Fanuc KAREL source: kb00020.KL

-- PROVISIONAL review KL for V1013-1; original PC SHA256 263743b7339b4aa91b7758d7d4a13bb68c8eefb6f044f5db318412e122d69ff7
-- Incomplete behavior may be omitted. Consult companion uncertainty JSON. Do not deploy.
PROGRAM KB00020
%NOLOCKGROUP
VAR
  P1 : INTEGER
  RESULT : STRING[80]
BEGIN
  -- UNRESOLVED_PC offsets 5-12; opcodes 9D,23
  -- UNRESOLVED_PC offsets 17-32; opcodes 27,22,76,75
  -- UNRESOLVED_PC offsets 37-41; opcodes 7F
END KB00020
